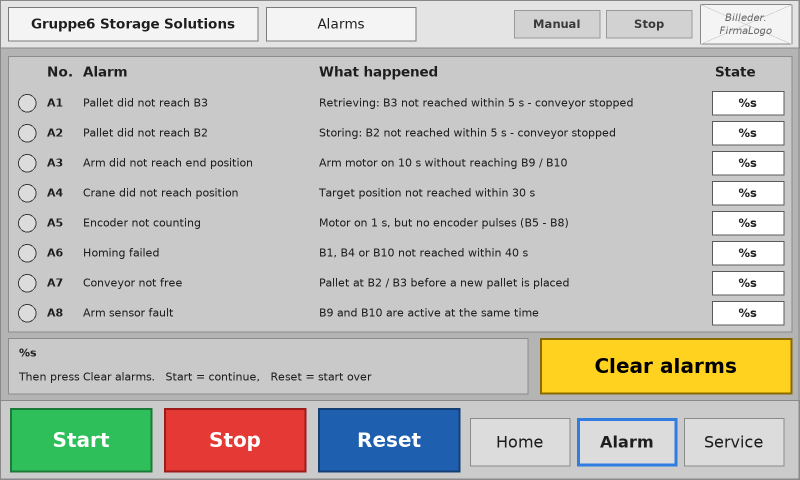
VISUALIZATION Alarm  // 800x480
    Rectangle (0,0 800x480)
    Rectangle (0,0 800x48)
    Rectangle (8,7 250x34), "Gruppe6 Storage Solutions"
    Rectangle (266,7 150x34), "Alarms"
    Rectangle (514,10 86x28), "Manual", colour toggle: MAIN.isManualMode
    Rectangle (606,10 86x28), "Stop", colour toggle: MAIN.isStop
    Image (700,4 92x40), image: Billeder.FirmaLogo
    Rectangle (0,400 800x80)
    RoundedRectangle (10,408 142x64), "Start"
        OnMouseUp: execute { MAIN.isStop := FALSE; }
    RoundedRectangle (164,408 142x64), "Stop"
        OnMouseUp: execute { MAIN.isStop := TRUE; }
    Rectangle (470,418 100x48), "Home"
        OnMouseUp: execute {
            MAIN.logoutRequest := TRUE;   // going to the Home page also logs out of the service page
        }
        OnMouseUp: change screen: Start
    Rectangle (684,418 100x48), "Service"
        OnMouseUp: change screen: Service
    Rectangle (577,418 100x48), "Alarm", colour toggle: MAIN.isAlarm
    Rectangle (8,56 784x276)
    Rectangle (44,60 34x24), "No."
    Rectangle (80,60 230x24), "Alarm"
    Rectangle (316,60 390x24), "What happened"
    Rectangle (712,60 72x24), "State"
    Ellipse (18,94 18x18), colour toggle: MAIN.alarmActive[1]
    Rectangle (44,90 34x26), "A1"
    Rectangle (80,90 230x26), "Pallet did not reach B3"
    Rectangle (316,90 390x26), "Retrieving: B3 not reached within 5 s - conveyor stopped"
    Rectangle (712,91 72x24), "%s", text variable: MAIN.alarmStateText[1], colour toggle: MAIN.alarmActive[1]
    Ellipse (18,124 18x18), colour toggle: MAIN.alarmActive[2]
    Rectangle (44,120 34x26), "A2"
    Rectangle (80,120 230x26), "Pallet did not reach B2"
    Rectangle (316,120 390x26), "Storing: B2 not reached within 5 s - conveyor stopped"
    Rectangle (712,121 72x24), "%s", text variable: MAIN.alarmStateText[2], colour toggle: MAIN.alarmActive[2]
    Ellipse (18,154 18x18), colour toggle: MAIN.alarmActive[3]
    Rectangle (44,150 34x26), "A3"
    Rectangle (80,150 230x26), "Arm did not reach end position"
    Rectangle (316,150 390x26), "Arm motor on 10 s without reaching B9 / B10"
    Rectangle (712,151 72x24), "%s", text variable: MAIN.alarmStateText[3], colour toggle: MAIN.alarmActive[3]
    Ellipse (18,184 18x18), colour toggle: MAIN.alarmActive[4]
    Rectangle (44,180 34x26), "A4"
    Rectangle (80,180 230x26), "Crane did not reach position"
    Rectangle (316,180 390x26), "Target position not reached within 30 s"
    Rectangle (712,181 72x24), "%s", text variable: MAIN.alarmStateText[4], colour toggle: MAIN.alarmActive[4]
    Ellipse (18,214 18x18), colour toggle: MAIN.alarmActive[5]
    Rectangle (44,210 34x26), "A5"
    Rectangle (80,210 230x26), "Encoder not counting"
    Rectangle (316,210 390x26), "Motor on 1 s, but no encoder pulses (B5 - B8)"
    Rectangle (712,211 72x24), "%s", text variable: MAIN.alarmStateText[5], colour toggle: MAIN.alarmActive[5]
    Ellipse (18,244 18x18), colour toggle: MAIN.alarmActive[6]
    Rectangle (44,240 34x26), "A6"
    Rectangle (80,240 230x26), "Homing failed"
    Rectangle (316,240 390x26), "B1, B4 or B10 not reached within 40 s"
    Rectangle (712,241 72x24), "%s", text variable: MAIN.alarmStateText[6], colour toggle: MAIN.alarmActive[6]
    Ellipse (18,274 18x18), colour toggle: MAIN.alarmActive[7]
    Rectangle (44,270 34x26), "A7"
    Rectangle (80,270 230x26), "Conveyor not free"
    Rectangle (316,270 390x26), "Pallet at B2 / B3 before a new pallet is placed"
    Rectangle (712,271 72x24), "%s", text variable: MAIN.alarmStateText[7], colour toggle: MAIN.alarmActive[7]
    Ellipse (18,304 18x18), colour toggle: MAIN.alarmActive[8]
    Rectangle (44,300 34x26), "A8"
    Rectangle (80,300 230x26), "Arm sensor fault"
    Rectangle (316,300 390x26), "B9 and B10 are active at the same time"
    Rectangle (712,301 72x24), "%s", text variable: MAIN.alarmStateText[8], colour toggle: MAIN.alarmActive[8]
    Rectangle (8,338 520x56)
    Rectangle (16,341 504x24), "%s", text variable: MAIN.alarmHelpText
    Rectangle (16,365 504x24), "Then press Clear alarms. Start = continue, Reset = start over"
    RoundedRectangle (540,338 252x56), "Clear alarms"
        OnMouseUp: execute {
            MAIN.alarmClearRequest := TRUE;   // clear all alarms
        }
    RoundedRectangle (318,408 142x64), "Reset"
        OnMouseUp: execute {
            MAIN.resetRequest := TRUE;   // everything back to Step_10, then homing
        }
END_VISUALIZATION

(* stored: Version 1.1.0.1, ProductVersion 3.1.4024.12
   Visu Alarm: Id {51597b5a-f402-4588-9aca-ebda3a23a9f6} *)
